Fanuc KAREL source: kt00266.KL

-- PROVISIONAL review KL for V770-1; original PC SHA256 9ae27d0fc5547d5c31850c197062d23a7c1182aebce7af6bb5dba4023680ecd1
-- Incomplete behavior may be omitted. Consult companion uncertainty JSON. Do not deploy.
PROGRAM KT00266
%NOLOCKGROUP
VAR
  S1 : STRING[80]
  S2 : STRING[80]
  OUT : BOOLEAN
BEGIN
  -- UNRESOLVED_PC offsets 5-14; opcodes 3F,75
  -- UNRESOLVED_PC offsets 19-28; opcodes 3F,75
  -- UNRESOLVED_PC offsets 33-42; opcodes 3F,75
  -- UNRESOLVED_PC offsets 47-56; opcodes 3F,75
  -- UNRESOLVED_PC offsets 61-80; opcodes 73,73,83,23
  -- UNRESOLVED_PC offsets 85-89; opcodes 7F
END KT00266
